(* IEC 61131-3 sources: SRCI_CLIENT_PLC/RobotLibrary/Library/POUs/Read/MC_ReadRobotSWLimits/Structures, 4 files *)

(* ---- ReadRobotSWLimitsOutCmd.st ---- *)
{attribute 'pack_mode' := '1'}
// -------------------------------------------------------------------------
//  SRCI Robot Library
// -------------------------------------------------------------------------
//
//  Object:      ReadRobotSWLimitsOutCmd
//  Author:      Thorsten Brach
//  Date:        2024-08-09
//
//  Description:
//
//
//  Copyright:
//    (C) 2024 Thorsten Brach. All rights reserved
//             Licensed under the MIT License.
//
//  Disclaimer:
//    This project is provided without any guarantee and can be used for
//    private and commercial purposes. Any use is at the user’s
//    own risk and responsibility.
//
// -------------------------------------------------------------------------
TYPE ReadRobotSWLimitsOutCmd :
STRUCT
  /// DLimits for joints and external axes according to Table 6-197.
  LimitValues        : SWLimits;
  /// The limits were changed on the RC since the last synchronization (ST-FIX F32: byte 106 of the response)
  DataChanged : BOOL;
END_STRUCT
END_TYPE

(* ---- ReadRobotSWLimitsParCmd.st ---- *)
{attribute 'pack_mode' := '1'}
// -------------------------------------------------------------------------
//  SRCI Robot Library
// -------------------------------------------------------------------------
//
//  Object:      ReadRobotSWLimitsParCmd
//  Author:      Thorsten Brach
//  Date:        2024-08-09
//
//  Description:
//
//
//  Copyright:
//    (C) 2024 Thorsten Brach. All rights reserved
//             Licensed under the MIT License.
//
//  Disclaimer:
//    This project is provided without any guarantee and can be used for
//    private and commercial purposes. Any use is at the user’s
//    own risk and responsibility.
//
// -------------------------------------------------------------------------
TYPE ReadRobotSWLimitsParCmd :
STRUCT
END_STRUCT
END_TYPE

(* ---- ReadRobotSWLimitsRecvData.st ---- *)
{attribute 'pack_mode' := '1'}
// -------------------------------------------------------------------------
//  SRCI Robot Library
// -------------------------------------------------------------------------
//
//  Object:      ReadRobotSWLimitsRecvData
//  Author:      Thorsten Brach
//  Date:        2024-08-09
//
//  Description:
//
//
//  Copyright:
//    (C) 2024 Thorsten Brach. All rights reserved
//             Licensed under the MIT License.
//
//  Disclaimer:
//    This project is provided without any guarantee and can be used for
//    private and commercial purposes. Any use is at the user’s
//    own risk and responsibility.
//
// -------------------------------------------------------------------------
TYPE ReadRobotSWLimitsRecvData EXTENDS RspHeader :
STRUCT
  /// DLimits for joints and external axes according to Table 6-197.
  LimitValues        : SWLimits;
  /// The status bit "DataChanged" represents the modification state
  DataChanged : BOOL;
END_STRUCT
END_TYPE

(* ---- ReadRobotSWLimitsSendData.st ---- *)
{attribute 'pack_mode' := '1'}
// -------------------------------------------------------------------------
//  SRCI Robot Library
// -------------------------------------------------------------------------
//
//  Object:      ReadRobotSWLimitsSendData
//  Author:      Thorsten Brach
//  Date:        2024-08-09
//
//  Description:
//
//
//  Copyright:
//    (C) 2024 Thorsten Brach. All rights reserved
//             Licensed under the MIT License.
//
//  Disclaimer:
//    This project is provided without any guarantee and can be used for
//    private and commercial purposes. Any use is at the user’s
//    own risk and responsibility.
//
// -------------------------------------------------------------------------
TYPE ReadRobotSWLimitsSendData EXTENDS CmdHeader:
STRUCT
END_STRUCT
END_TYPE
